Fanuc KAREL source: KT00991.KL

PROGRAM KT00991
%NOLOCKGROUP
VAR
  P1: POSITION
  P2: POSITION
  X: REAL
  Y: REAL
  Z: REAL
  W: REAL
  P: REAL
  R: REAL
  CFG: CONFIG
BEGIN
  UNPOS(P1, X, Y, Z, W, P, R, CFG)
END KT00991
